// CFC twin of T_SafeInputPair_Tests: the same tests drawn as CFC diagrams, the way a TwinSAFE project is authored.
    FUNCTION_BLOCK T_SafeInputPair_Tests_CFC EXTENDS T_SafeCfcTestSuite
    VAR
    // Test_InactivePairNeverRequestsSafeState
    pair_1 : T_SafeInputPair;
    // Test_BreakContactRequestsSafeStateOnZero
    pair_2 : T_SafeInputPair;
    // Test_MakeContactRequestsSafeStateOnOne
    pair_3 : T_SafeInputPair;
    // Test_TwoChannelRequestsSafeStateIfEitherChannelLow
    pair_4 : T_SafeInputPair;
    // Test_DiscrepancyErrorAfterTimeoutAndResetAfterSafeInputs
    pair_5 : T_SafeInputPair;
    t1_5 : TON;
    t2_5 : TON;
    trig1_5 : R_TRIG;
    trig2_5 : R_TRIG;
END_VAR

Test_InactivePairNeverRequestsSafeState();
Test_BreakContactRequestsSafeStateOnZero();
Test_MakeContactRequestsSafeStateOnOne();
Test_TwoChannelRequestsSafeStateIfEitherChannelLow();
Test_DiscrepancyErrorAfterTimeoutAndResetAfterSafeInputs();

METHOD PRIVATE Test_InactivePairNeverRequestsSafeState
// note: this text did not pass the execution check against the stored diagram
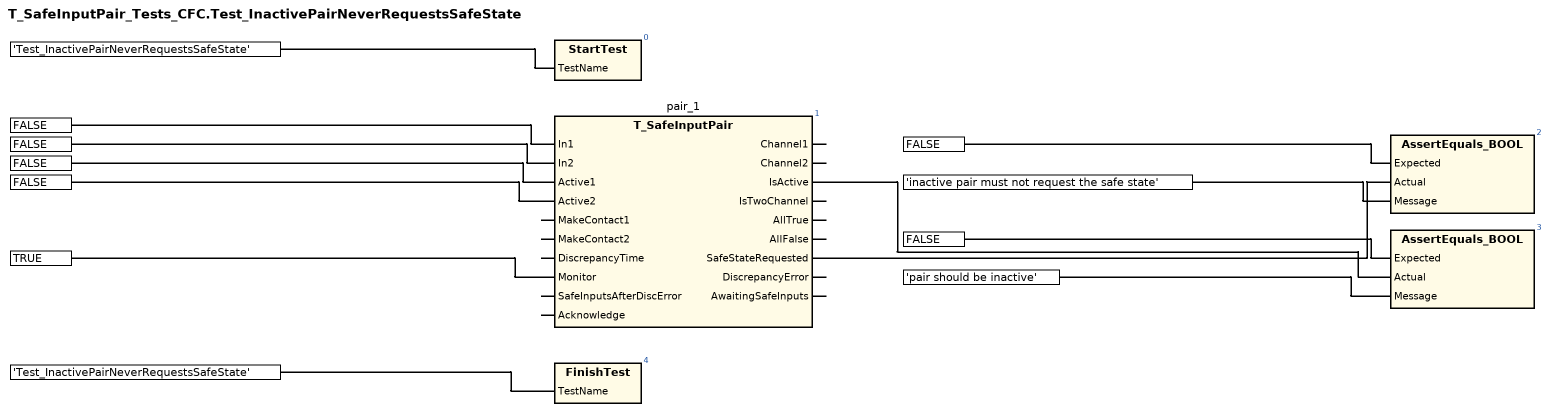
StartTest(TestName := 'Test_InactivePairNeverRequestsSafeState');
pair_1(In1 := FALSE, In2 := FALSE, Active1 := FALSE, Active2 := FALSE, Monitor := TRUE); // T_SafeInputPair
AssertEquals_BOOL(Expected := FALSE, Actual := pair_1.SafeStateRequested, Message := 'inactive pair must not request the safe state');
AssertEquals_BOOL(Expected := FALSE, Actual := pair_1.IsActive, Message := 'pair should be inactive');
FinishTest(TestName := 'Test_InactivePairNeverRequestsSafeState');
END_METHOD

METHOD PRIVATE Test_BreakContactRequestsSafeStateOnZero
// note: this text did not pass the execution check against the stored diagram
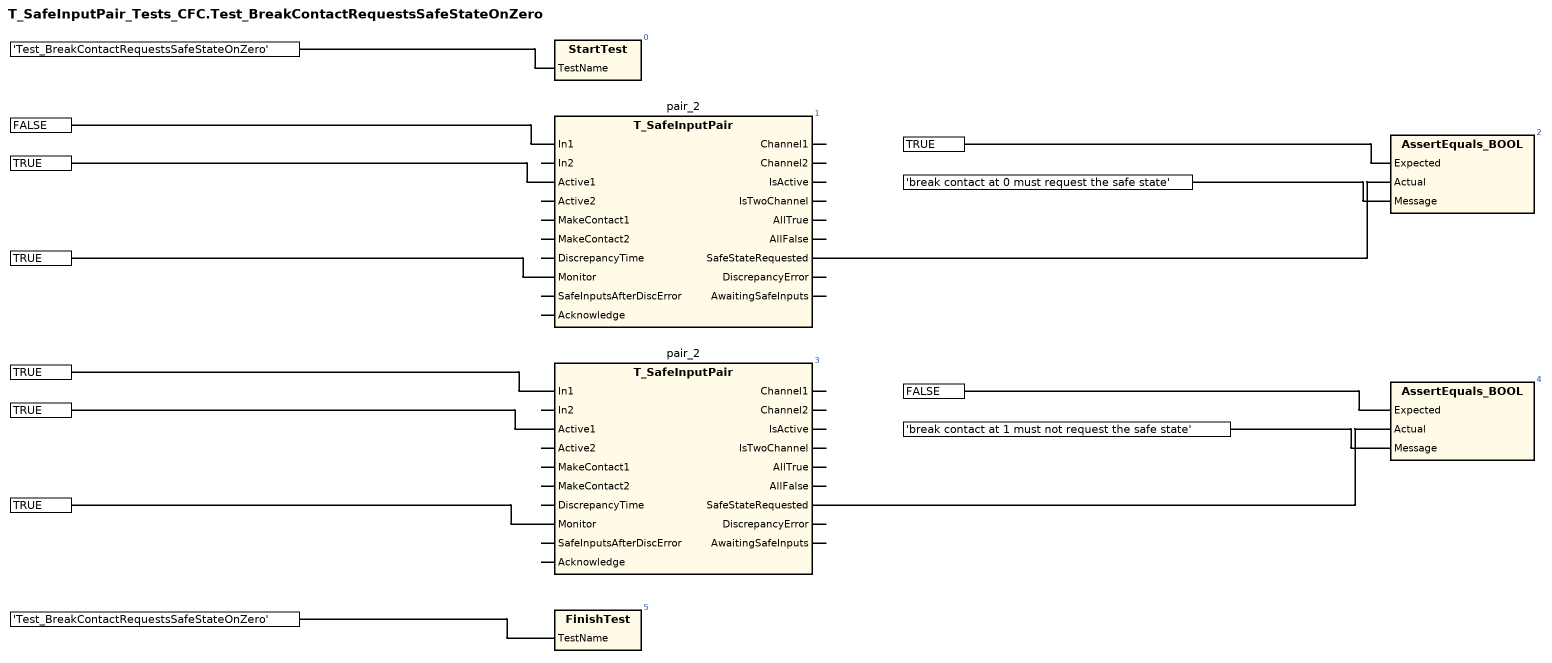
StartTest(TestName := 'Test_BreakContactRequestsSafeStateOnZero');
pair_2(In1 := FALSE, Active1 := TRUE, Monitor := TRUE); // T_SafeInputPair
AssertEquals_BOOL(Expected := TRUE, Actual := pair_2.SafeStateRequested, Message := 'break contact at 0 must request the safe state');
pair_2(In1 := TRUE, Active1 := TRUE, Monitor := TRUE); // T_SafeInputPair
AssertEquals_BOOL(Expected := FALSE, Actual := pair_2.SafeStateRequested, Message := 'break contact at 1 must not request the safe state');
FinishTest(TestName := 'Test_BreakContactRequestsSafeStateOnZero');
END_METHOD

METHOD PRIVATE Test_MakeContactRequestsSafeStateOnOne
// note: this text did not pass the execution check against the stored diagram
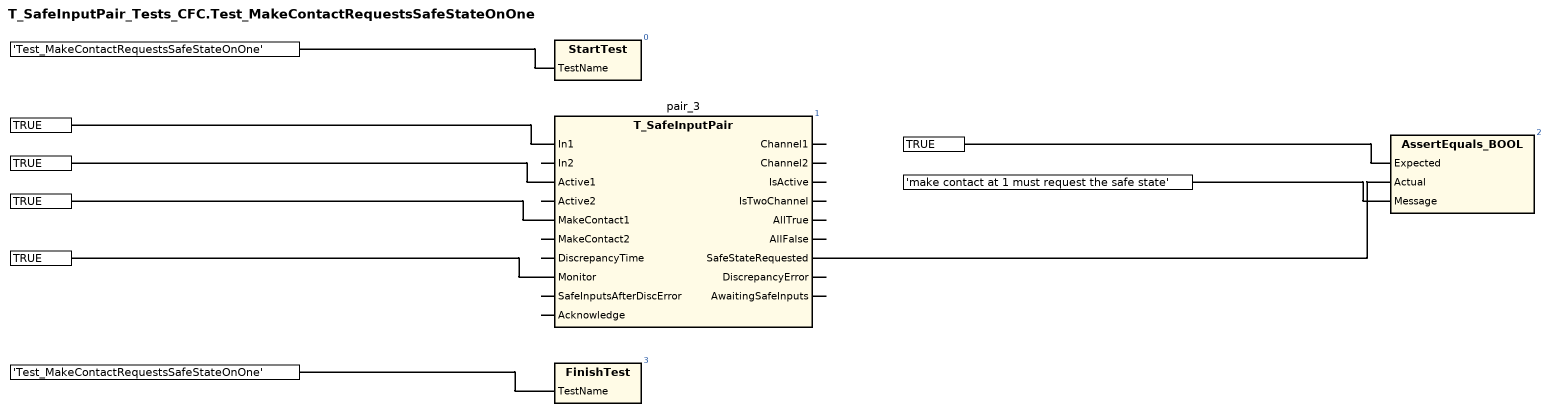
StartTest(TestName := 'Test_MakeContactRequestsSafeStateOnOne');
pair_3(In1 := TRUE, Active1 := TRUE, MakeContact1 := TRUE, Monitor := TRUE); // T_SafeInputPair
AssertEquals_BOOL(Expected := TRUE, Actual := pair_3.SafeStateRequested, Message := 'make contact at 1 must request the safe state');
FinishTest(TestName := 'Test_MakeContactRequestsSafeStateOnOne');
END_METHOD

METHOD PRIVATE Test_TwoChannelRequestsSafeStateIfEitherChannelLow
// note: this text did not pass the execution check against the stored diagram
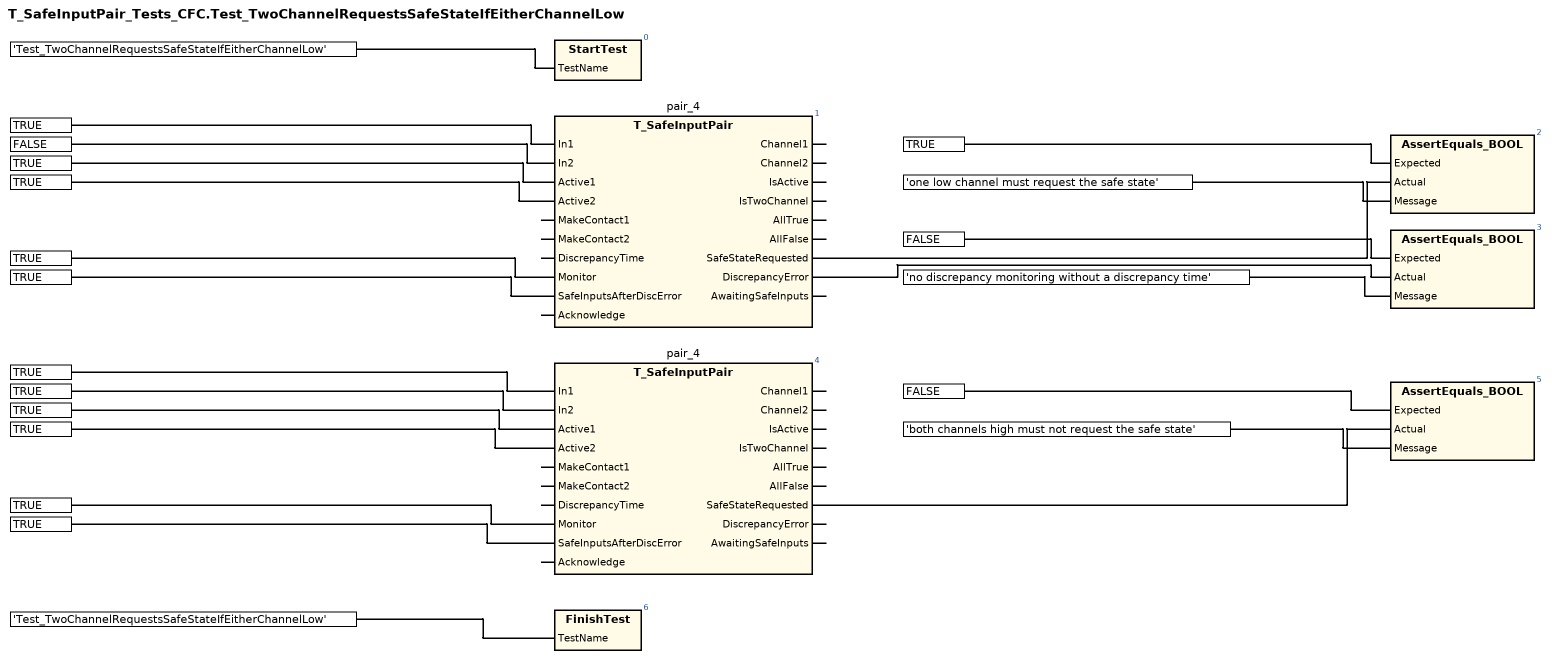
StartTest(TestName := 'Test_TwoChannelRequestsSafeStateIfEitherChannelLow');
pair_4(
    In1 := TRUE,
    In2 := FALSE,
    Active1 := TRUE,
    Active2 := TRUE,
    Monitor := TRUE,
    SafeInputsAfterDiscError := TRUE); // T_SafeInputPair
AssertEquals_BOOL(Expected := TRUE, Actual := pair_4.SafeStateRequested, Message := 'one low channel must request the safe state');
AssertEquals_BOOL(Expected := FALSE, Actual := pair_4.DiscrepancyError, Message := 'no discrepancy monitoring without a discrepancy time');
pair_4(
    In1 := TRUE,
    In2 := TRUE,
    Active1 := TRUE,
    Active2 := TRUE,
    Monitor := TRUE,
    SafeInputsAfterDiscError := TRUE); // T_SafeInputPair
AssertEquals_BOOL(Expected := FALSE, Actual := pair_4.SafeStateRequested, Message := 'both channels high must not request the safe state');
FinishTest(TestName := 'Test_TwoChannelRequestsSafeStateIfEitherChannelLow');
END_METHOD

METHOD PRIVATE Test_DiscrepancyErrorAfterTimeoutAndResetAfterSafeInputs
// note: this text did not pass the execution check against the stored diagram
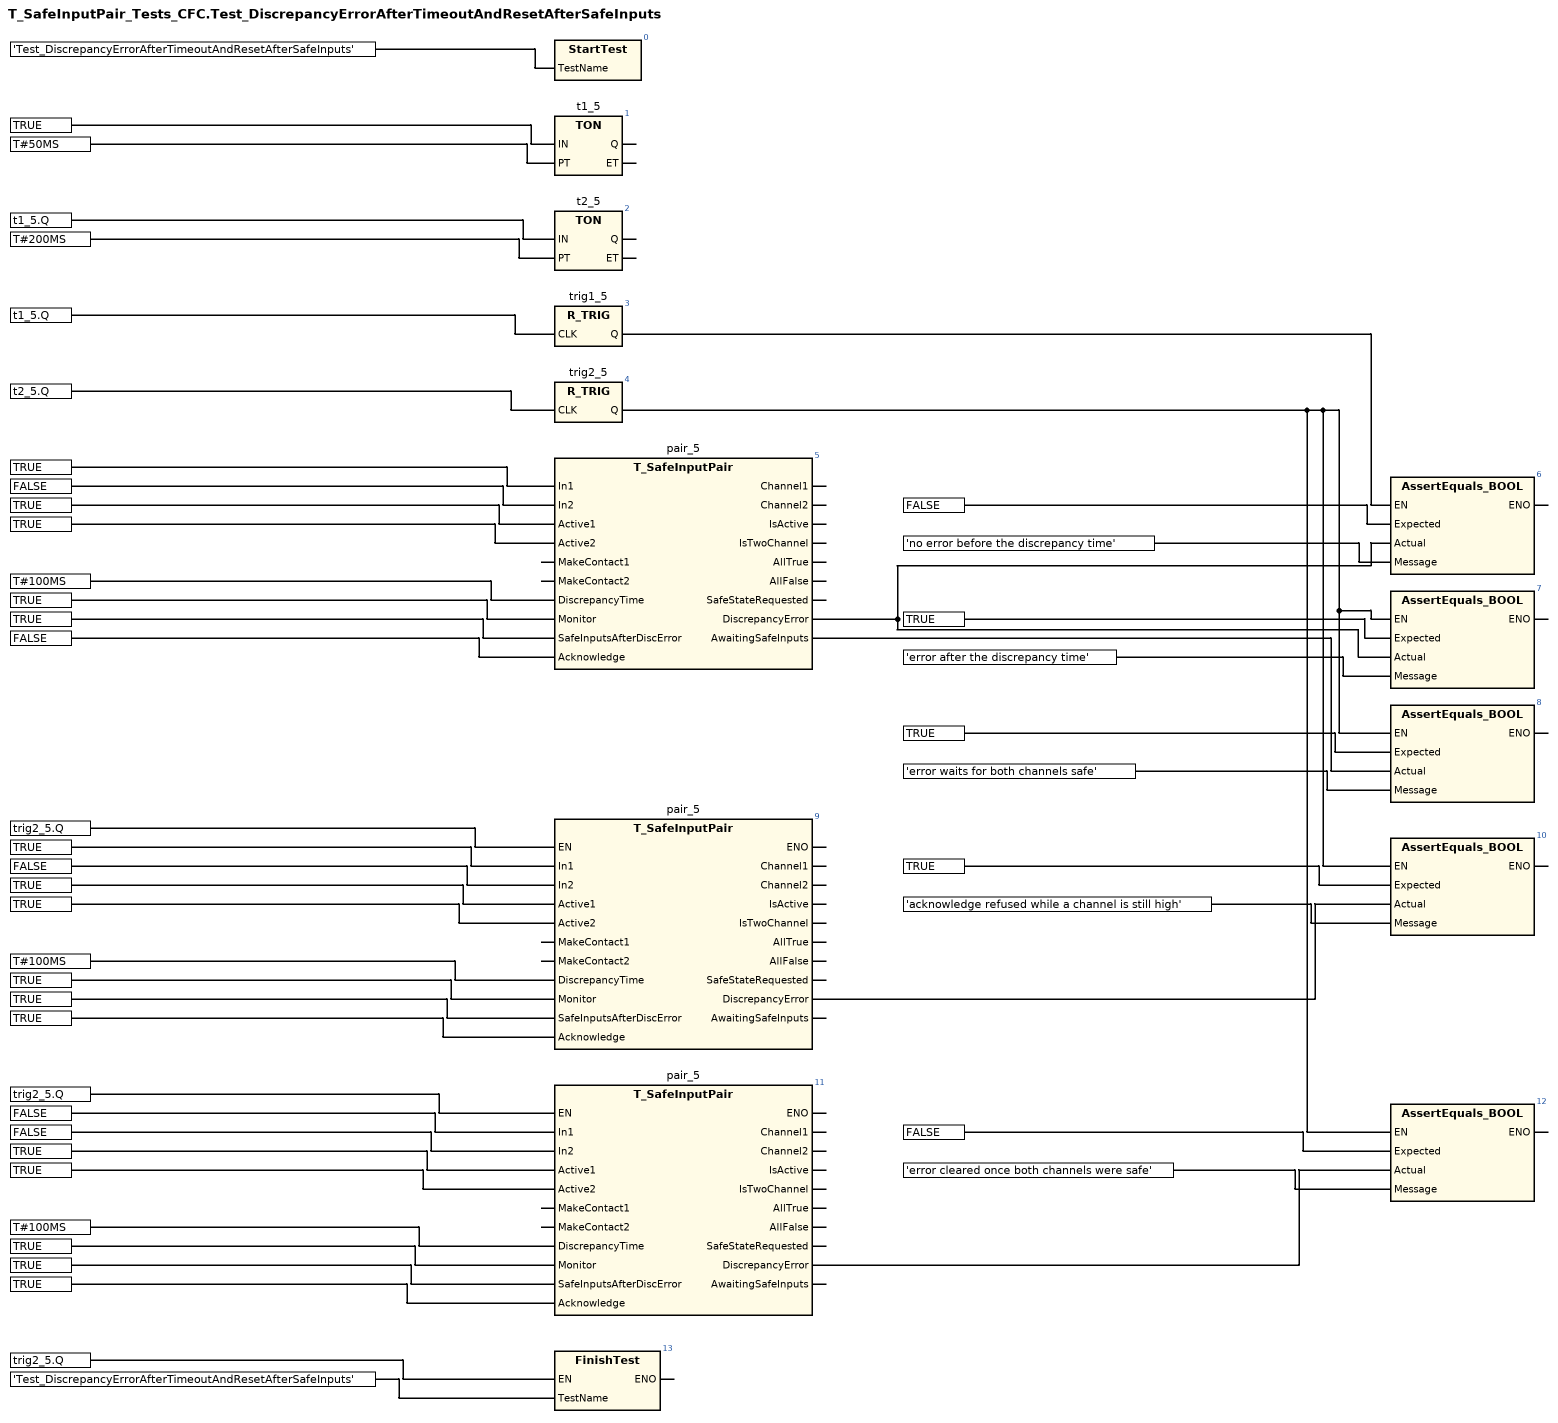
StartTest(TestName := 'Test_DiscrepancyErrorAfterTimeoutAndResetAfterSafeInputs');
t1_5(IN := TRUE, PT := T#50MS); // TON
t2_5(IN := t1_5.Q, PT := T#200MS); // TON
trig1_5(CLK := t1_5.Q); // R_TRIG
trig2_5(CLK := t2_5.Q); // R_TRIG
pair_5(
    In1 := TRUE,
    In2 := FALSE,
    Active1 := TRUE,
    Active2 := TRUE,
    DiscrepancyTime := T#100MS,
    Monitor := TRUE,
    SafeInputsAfterDiscError := TRUE,
    Acknowledge := FALSE); // T_SafeInputPair
IF trig1_5.Q THEN AssertEquals_BOOL(Expected := FALSE, Actual := pair_5.DiscrepancyError, Message := 'no error before the discrepancy time'); END_IF
IF trig2_5.Q THEN AssertEquals_BOOL(Expected := TRUE, Actual := pair_5.DiscrepancyError, Message := 'error after the discrepancy time'); END_IF
IF trig2_5.Q THEN AssertEquals_BOOL(Expected := TRUE, Actual := pair_5.AwaitingSafeInputs, Message := 'error waits for both channels safe'); END_IF
IF trig2_5.Q THEN
    pair_5(
        In1 := TRUE,
        In2 := FALSE,
        Active1 := TRUE,
        Active2 := TRUE,
        DiscrepancyTime := T#100MS,
        Monitor := TRUE,
        SafeInputsAfterDiscError := TRUE,
        Acknowledge := TRUE); // T_SafeInputPair
END_IF
IF trig2_5.Q THEN AssertEquals_BOOL(Expected := TRUE, Actual := pair_5.DiscrepancyError, Message := 'acknowledge refused while a channel is still high'); END_IF
IF trig2_5.Q THEN
    pair_5(
        In1 := FALSE,
        In2 := FALSE,
        Active1 := TRUE,
        Active2 := TRUE,
        DiscrepancyTime := T#100MS,
        Monitor := TRUE,
        SafeInputsAfterDiscError := TRUE,
        Acknowledge := TRUE); // T_SafeInputPair
END_IF
IF trig2_5.Q THEN AssertEquals_BOOL(Expected := FALSE, Actual := pair_5.DiscrepancyError, Message := 'error cleared once both channels were safe'); END_IF
IF trig2_5.Q THEN FinishTest(TestName := 'Test_DiscrepancyErrorAfterTimeoutAndResetAfterSafeInputs'); END_IF
END_METHOD

END_FUNCTION_BLOCK

(* stored: Version 1.1.0.1, ProductVersion 3.1.4026.22
   POU T_SafeInputPair_Tests_CFC: Id {cc86fd5c-5f7c-5925-9bca-64feebc6c714}, SpecialFunc None
   Method Test_InactivePairNeverRequestsSafeState: Id {53252cd9-dd48-5ef5-a58d-9217164443f1}
   Method Test_BreakContactRequestsSafeStateOnZero: Id {17ef0ab5-9c27-513b-a8e8-9861b19ae44a}
   Method Test_MakeContactRequestsSafeStateOnOne: Id {60d845e1-8f2a-5454-a667-f7465ef02b1a}
   Method Test_TwoChannelRequestsSafeStateIfEitherChannelLow: Id {9c9f94fd-2e4a-5c19-bc3c-5d6df0516d5b}
   Method Test_DiscrepancyErrorAfterTimeoutAndResetAfterSafeInputs: Id {e10d3a81-3aff-5101-882e-400211d05bc0} *)
